Staubli VAL3: simulate.pgx

program simulate()
begin
end
